(* IEC 61131-3 sources: Test-Git_ESME26/TestProgettoESME_26.fbsproj/PacDriveLib Migration/Motion/Control/PDL_FB_DriveEnable.fb.st^, 3 files *)

(* ---- Init.meth.st ---- *)
{attribute 'hide'}
METHOD PRIVATE Init : BOOL
VAR_INPUT
END_VAR

Init := FALSE;

IF i_ifDrive <> 0 THEN
	fbStop.Axis := i_ifDrive;
	fbPower.Axis := i_ifDrive;
	fbReset.Axis := i_ifDrive;
ELSE
	SetDiagOutput(	i_etDiag	:= GD.ET_Diag.InputParameterInvalid,
					i_etDiagExt := PDL_ET_DiagExt.DriveInvalid,
					i_sMsg		:= 'i_ifDrive - Invalid Interface');
	RETURN;
END_IF

xSuccess := __QUERYINTERFACE(i_ifDrive, ifGetParentDevice);
IF NOT xSuccess THEN
	SetDiagOutput(	i_etDiag	:= GD.ET_Diag.InputParameterInvalid,
					i_etDiagExt := PDL_ET_DiagExt.DriveInvalid,
					i_sMsg		:= 'i_ifDrive - DTSI.IF_GetParentDevice not implemented');
	RETURN;
END_IF

ifDeviceAccess := ifGetParentDevice.GetParentDevice();
xSuccess := __QUERYINTERFACE(ifDeviceAccess, ifDiagnosticAccess);
IF xSuccess THEN
	ifDiagnostic := ifDiagnosticAccess.Diagnostic;
ELSE
	SetDiagOutput(	i_etDiag	:= GD.ET_Diag.InputParameterInvalid,
					i_etDiagExt := PDL_ET_DiagExt.DriveInvalid,
					i_sMsg		:= 'i_ifDrive - UFMPLCI.IF_DiagnosticAccess not implemented');
	RETURN;
END_IF

xSuccess := __QUERYINTERFACE(ifDeviceAccess, ifDriveConfigAccess);
IF xSuccess THEN
	ifDriveConfig := ifDriveConfigAccess.DriveConfig;
ELSE
	SetDiagOutput(	i_etDiag	:= GD.ET_Diag.InputParameterInvalid,
					i_etDiagExt := PDL_ET_DiagExt.DriveInvalid,
					i_sMsg		:= 'i_ifDrive - DDI.IF_DriveConfigAccess not implemented');
	RETURN;
END_IF

xSuccess := __QUERYINTERFACE(ifDeviceAccess, ifDrivePowerSupplyAccess);
IF xSuccess THEN
	ifDrivePowerSupply := ifDrivePowerSupplyAccess.DrivePowerSupply;
ELSE
	SetDiagOutput(	i_etDiag	:= GD.ET_Diag.InputParameterInvalid,
					i_etDiagExt := PDL_ET_DiagExt.DriveInvalid,
					i_sMsg		:= 'i_ifDrive - DDI.IF_DrivePowerSupplyAccess not implemented');
	RETURN;
END_IF

xSuccess := __QUERYINTERFACE(ifDeviceAccess, ifWorkingModeAccess);
IF xSuccess THEN
	ifWorkingMode := ifWorkingModeAccess.WorkingMode;
ELSE
	SetDiagOutput(	i_etDiag	:= GD.ET_Diag.InputParameterInvalid,
					i_etDiagExt := PDL_ET_DiagExt.DriveInvalid,
					i_sMsg		:= 'i_ifDrive - DDI.IF_DrivePowerSupplyAccess not implemented');
	RETURN;
END_IF

IF ifWorkingMode.ActualState = CFDI.ET_WorkingState.Physical THEN
	ifPowerSupplyDevice := ifDrivePowerSupply.GetDevice();
	xSuccess := __QUERYINTERFACE(ifPowerSupplyDevice, ifPowerSupplyAccess);
	IF xSuccess THEN
		ifPowerSupply := ifPowerSupplyAccess.PowerSupply;
	ELSE
		SetDiagOutput(	i_etDiag	:= GD.ET_Diag.InputParameterInvalid,
						i_etDiagExt := PDL_ET_DiagExt.DriveInvalid,
						i_sMsg		:= 'i_ifDrive - DDI.IF_PowerSupplyAccess not implemented');
		RETURN;
	END_IF

	xSuccess := __QUERYINTERFACE(ifPowerSupplyDevice, ifPowerSupplyDiagnosticAccess);
	IF xSuccess THEN
		ifPowerSupplyDiagnostic := ifPowerSupplyDiagnosticAccess.Diagnostic;
	ELSE
		SetDiagOutput(	i_etDiag	:= GD.ET_Diag.InputParameterInvalid,
						i_etDiagExt := PDL_ET_DiagExt.DriveInvalid,
						i_sMsg		:= 'PowerSupply - UFMPLCI.IF_DiagnosticAccess not implemented');
		RETURN;
	END_IF
	xDriveIsReal := TRUE;
	Init := TRUE;
ELSE
	xDriveIsReal := FALSE;
	Init := TRUE;
END_IF

xSuccess := __QUERYINTERFACE(ifDeviceAccess, ifDeviceTreeObjectAccess);
IF xSuccess THEN
	sDriveName := ifDeviceTreeObjectAccess.DeviceTreeObject.Name;
ELSE
	sDriveName := 'Axis';
END_IF

(* ---- RegisterLoggerPoint.meth.st ---- *)
METHOD PUBLIC RegisterLoggerPoint
VAR_INPUT
	i_ifParent		: APL.IF_LoggerPoint;
	i_sName			: STRING[80];
END_VAR
VAR_OUTPUT
	q_etDiag		: GD.ET_Diag := GD.ET_Diag.Ok;
	q_etDiagExt		: PDL_ET_DiagExt := PDL_ET_DiagExt.Ok;
END_VAR
VAR
	etDiagBuffer		: GD.ET_Diag;
	etDiagExtBufferAPL	: APL.ET_DiagExt;
END_VAR

THIS^.fbLoggerPoint.RegisterLoggerPoint(	i_ifParent		:= i_ifParent,
											i_sName			:= i_sName,
											i_sType			:= 'FB_DriveEnable',
											i_sSource		:= 'PDL',
											q_etDiag		=> etDiagBuffer,
											q_etDiagExt		=> etDiagExtBufferAPL);
IF (etDiagBuffer <> GD.ET_Diag.Ok) THEN
	CASE etDiagExtBufferAPL OF
		APL.ET_DiagExt.ParentInvalid:
			q_etDiag := GD.ET_Diag.InputParameterInvalid;
			q_etDiagExt := PDL_ET_DiagExt.ParentInvalid;

		APL.ET_DiagExt.ParentNotRegistered:
			q_etDiag := GD.ET_Diag.InputParameterInvalid;
			q_etDiagExt := PDL_ET_DiagExt.ParentNotRegistered;

		APL.ET_DiagExt.MaxNumberOfLoggerPointsExeeded:
			q_etDiag := GD.ET_Diag.InputParameterInvalid;
			q_etDiagExt := PDL_ET_DiagExt.MaxNumberOfLoggerPointsExeeded;

	ELSE
		q_etDiag := GD.ET_Diag.UnexpectedProgramBehavior;
		q_etdiagExt := PDL_ET_DiagExt.UnexpectedDiagExt;
	END_CASE
END_IF

(* ---- SetDiagOutput.meth.st ---- *)
{attribute 'hide'}
METHOD SetDiagOutput : BOOL
VAR_INPUT
	i_etDiag	: GD.ET_Diag;
	i_etDiagExt	: PDL_ET_DiagExt;
	i_sMsg		: STRING[80];
END_VAR
VAR
END_VAR

IF i_etDiag <> GD.ET_Diag.Ok THEN
	q_xReady := FALSE;
END_IF

IF q_etDiag = GD.ET_Diag.OK OR i_etDiagExt = PDL_ET_DiagExt.Disabled THEN
	q_etDiag := i_etDiag;
	q_etDiagExt := i_etDiagExt;
	q_sMsg := i_sMsg;

	IF(i_etDiag = GD.ET_Diag.Ok) AND (THIS^.fbLoggerPoint.etLogLevel >= APL.ET_LogLevel.StatusMessage) THEN
		THIS^.fbLoggerPoint.AddLogEntry(	i_etLogLevel	:= APL.ET_LogLevel.StatusMessage,
											i_etDiag		:= q_etDiag,
											i_udiDiagExt	:= q_etDiagExt,
											i_sMessage		:= SE_CTBX.FC_MultiConcat(	i_sString1	:= Standard.CONCAT('ET_Diag: ', GD.FC_EtDiagToString(q_etDiag)),
																						i_sString2	:= Standard.CONCAT(' ET_DiagExt: ', PDL_FC_EtDiagExtToString(q_etDiagExt)),
																						i_sString3	:= Standard.CONCAT(' sMsg: ', q_sMsg),
																						i_sString4	:= '')
											);
	ELSIF(i_etDiag = GD.ET_Diag.UnexpectedProgramBehavior) AND (THIS^.fbLoggerPoint.etLogLevel >= APL.ET_LogLevel.CriticalException) THEN
		THIS^.fbLoggerPoint.AddLogEntry(	i_etLogLevel	:= APL.ET_LogLevel.CriticalException,
											i_etDiag		:= q_etDiag,
											i_udiDiagExt	:= q_etDiagExt,
											i_sMessage		:= SE_CTBX.FC_MultiConcat(	i_sString1	:= Standard.CONCAT('ET_Diag: ', GD.FC_EtDiagToString(q_etDiag)),
																						i_sString2	:= Standard.CONCAT(' ET_DiagExt: ', PDL_FC_EtDiagExtToString(q_etDiagExt)),
																						i_sString3	:= Standard.CONCAT(' sMsg: ', q_sMsg),
																						i_sString4	:= '')
											);
	ELSIF(i_etDiag <> GD.ET_Diag.Ok) AND (THIS^.fbLoggerPoint.etLogLevel >= APL.ET_LogLevel.Exception) THEN
		THIS^.fbLoggerPoint.AddLogEntry(	i_etLogLevel	:= APL.ET_LogLevel.Exception,
											i_etDiag		:= q_etDiag,
											i_udiDiagExt	:= q_etDiagExt,
											i_sMessage		:= SE_CTBX.FC_MultiConcat(	i_sString1	:= Standard.CONCAT('ET_Diag: ', GD.FC_EtDiagToString(q_etDiag)),
																				i_sString2	:= Standard.CONCAT(' ET_DiagExt: ', PDL_FC_EtDiagExtToString(q_etDiagExt)),
																				i_sString3	:= Standard.CONCAT(' sMsg: ', q_sMsg),
																				i_sString4	:= '')
											);
	END_IF
END_IF
